// TIA Portal V19 export
FUNCTION_BLOCK "ULTRACHILLED_SKIDS"   // FB17, LAD
{ S7_Optimized_Access := 'TRUE' }
// stored: MemoryReserve 100, SetENOAutomatically false
   VAR_INPUT
      TEMP_SP : Real;
      START : Bool;
      STOP : Bool;
      AUTO : Bool;
      EMG : Bool;
      FS_HE_INLET : Bool;
      FS_HE_OUTLET : Bool;
      MGLT_LSP : Real;
      HOLD_RESUME : Bool;
      TT01_fault : Bool;
      TT02_fault : Bool;
      TT03_fault : Bool;
      TT04_fault : Bool;
      MGLT_FAULT : Bool;
      PUMP_1RPM : Real;
      "PUMP_1RPM SP" : Real;
      "PUMP_2 RPM" : Real;
      "PUMP_2 RPM SP" : Real;
      HEADER_PSP : Real;
      HEADER_PRESSURE_PV : Real;
      TEMP_PV : Real;
      MGLT_PV : Real;
   END_VAR
   VAR_OUTPUT
      PUMP_1_CMD : Bool;
      PUMP_2_CMD : Bool;
      RUNNING : Bool;
      UCH_BUXV1501_CMD : Bool;
      PUMP_1_FAULTY : Bool;
      PUMP_2_FAULTY : Bool;
   END_VAR
   VAR
      "STEP" : Int;
      ALL_OK : Bool;
      IEC_Timer_0_Instance { S7_SetPoint := 'True'} : TP_TIME;
      P_TRIG_1 { S7_SetPoint := 'True'} : Bool;
      P_TRIG_2 : Bool;
      P_TRIG_3 : Bool;
      P_TRIG_4 : Bool;
      P_TRIG_5 : Bool;
      P_TRIG_6 : Bool;
      P_TRIG_7 : Bool;
      P_TRIG_8 : Bool;
   END_VAR
   VAR_TEMP   // added for the SCL form of the ladder/FBD networks
      _w1 : Bool;
      _w2 : Bool;
      _w3 : Bool;
      _w4 : Bool;
   END_VAR
BEGIN

REGION Network 1: PRECHECK
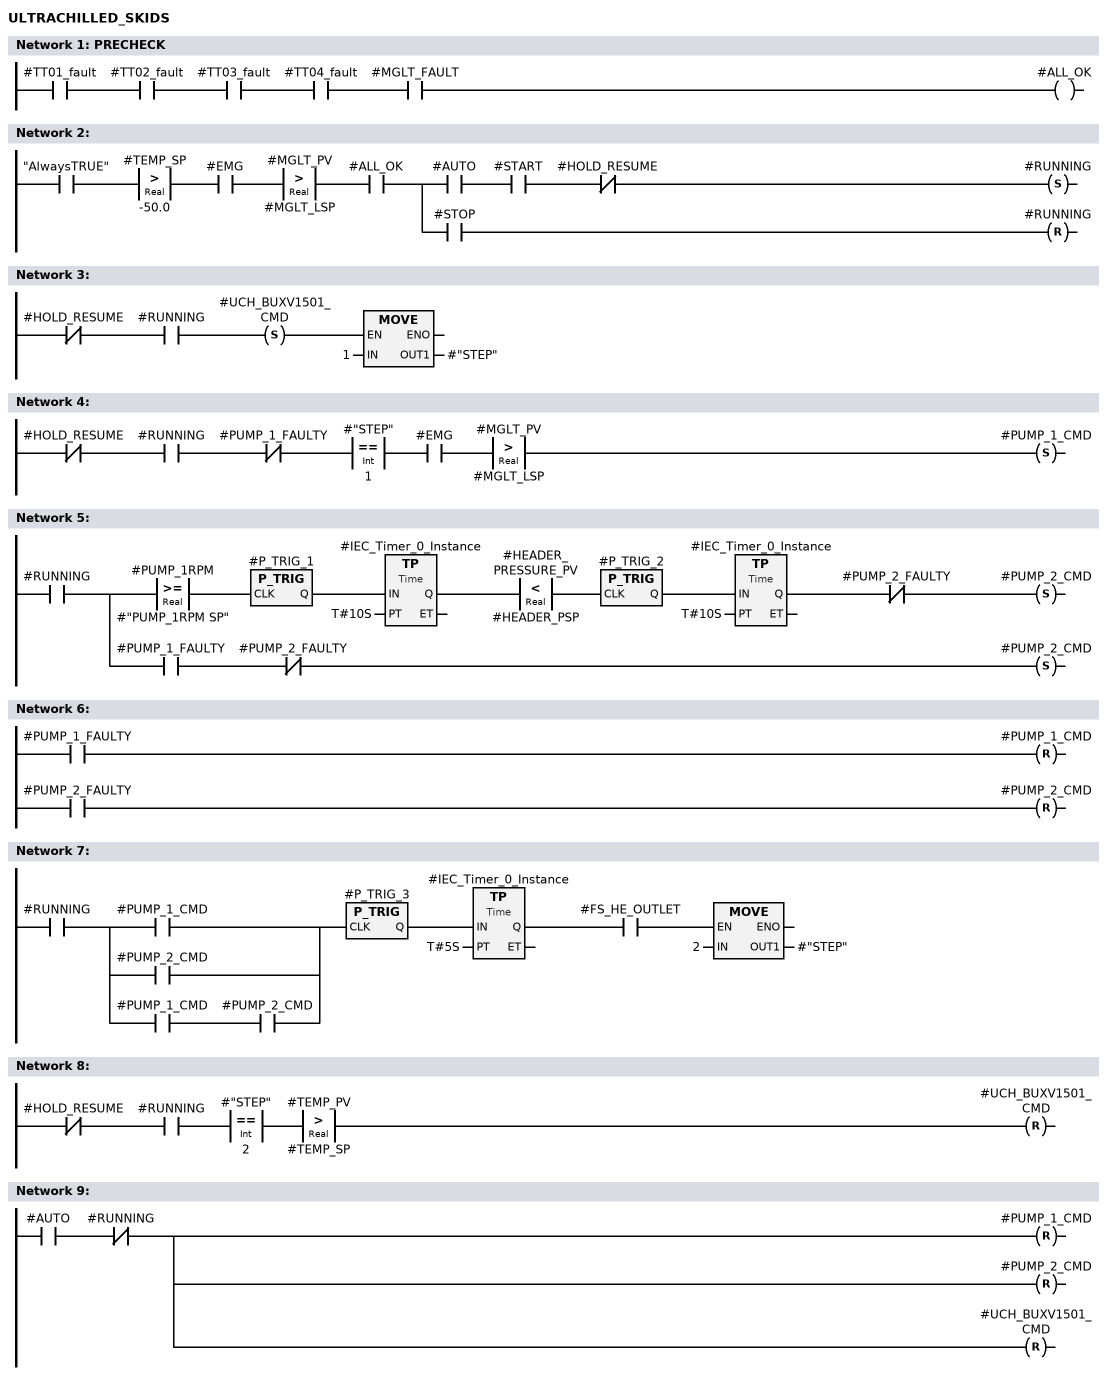
   RUNG wire#powerrail
      Contact( #TT01_fault )
      Contact( #TT02_fault )
      Contact( #TT03_fault )
      Contact( #TT04_fault )
      Contact( #MGLT_FAULT )
      Coil( #ALL_OK )
   END_RUNG
   // the same network as SCL:
   #ALL_OK := #TT01_fault AND #TT02_fault AND #TT03_fault AND #TT04_fault AND #MGLT_FAULT;
END_REGION

REGION Network 2
   RUNG wire#powerrail
      Contact( "AlwaysTRUE" )
      { S7_Templates := "SrcType := Real" } GT_Contact(in1 := #TEMP_SP, in2 := -50.0)
      Contact( #EMG )
      { S7_Templates := "SrcType := Real" } GT_Contact(in1 := #MGLT_PV, in2 := #MGLT_LSP)
      Contact( #ALL_OK )
      wire#w1
      Contact( #AUTO )
      Contact( #START )
      I_Contact( #HOLD_RESUME )
      S_Coil( #RUNNING )
   END_RUNG
   RUNG wire#w1
      Contact( #STOP )
      R_Coil( #RUNNING )
   END_RUNG
   // the same network as SCL:
   #_w1 := "AlwaysTRUE" AND (#TEMP_SP > (-50.0)) AND #EMG AND (#MGLT_PV > #MGLT_LSP) AND #ALL_OK;
   IF #_w1 AND #AUTO AND #START AND NOT #HOLD_RESUME THEN #RUNNING := TRUE; END_IF;
   IF #_w1 AND #STOP THEN #RUNNING := FALSE; END_IF;
END_REGION

REGION Network 3
   RUNG wire#powerrail
      I_Contact( #HOLD_RESUME )
      Contact( #RUNNING )
      S_Coil( #UCH_BUXV1501_CMD )
      Move(in := 1, out1 => #"STEP")
   END_RUNG
   // the same network as SCL:
   IF NOT #HOLD_RESUME AND #RUNNING THEN
       #UCH_BUXV1501_CMD := TRUE;
       #"STEP" := 1;
   END_IF;
END_REGION

REGION Network 4
   RUNG wire#powerrail
      I_Contact( #HOLD_RESUME )
      Contact( #RUNNING )
      I_Contact( #PUMP_1_FAULTY )
      { S7_Templates := "SrcType := Int" } EQ_Contact(in1 := #"STEP", in2 := 1)
      Contact( #EMG )
      { S7_Templates := "SrcType := Real" } GT_Contact(in1 := #MGLT_PV, in2 := #MGLT_LSP)
      S_Coil( #PUMP_1_CMD )
   END_RUNG
   // the same network as SCL:
   IF NOT #HOLD_RESUME AND #RUNNING AND NOT #PUMP_1_FAULTY AND (#"STEP" = 1) AND #EMG AND (#MGLT_PV > #MGLT_LSP) THEN
       #PUMP_1_CMD := TRUE;
   END_IF;
END_REGION

REGION Network 5
   RUNG wire#powerrail
      Contact( #RUNNING )
      wire#w1
      { S7_Templates := "SrcType := Real" } GE_Contact(in1 := #PUMP_1RPM, in2 := #"PUMP_1RPM SP")
      P_Trig( #P_TRIG_1 )
      { S7_Templates := "time_type := Time" } #IEC_Timer_0_Instance.TP(pt := T#10S, et =>)
      { S7_Templates := "SrcType := Real" } LT_Contact(in1 := #HEADER_PRESSURE_PV, in2 := #HEADER_PSP)
      P_Trig( #P_TRIG_2 )
      { S7_Templates := "time_type := Time" } #IEC_Timer_0_Instance.TP(pt := T#10S, et =>)
      I_Contact( #PUMP_2_FAULTY )
      S_Coil( #PUMP_2_CMD )
   END_RUNG
   RUNG wire#w1
      Contact( #PUMP_1_FAULTY )
      I_Contact( #PUMP_2_FAULTY )
      S_Coil( #PUMP_2_CMD )
   END_RUNG
   // the same network as SCL:
   #_w1 := #RUNNING AND (#PUMP_1RPM >= #"PUMP_1RPM SP");
   #_w2 := #_w1 AND NOT #P_TRIG_1;   // rising edge
   #P_TRIG_1 := #_w1;
   #IEC_Timer_0_Instance(IN := #_w2, PT := T#10S);   // TP
   #_w3 := #IEC_Timer_0_Instance.Q AND (#HEADER_PRESSURE_PV < #HEADER_PSP);
   #_w4 := #_w3 AND NOT #P_TRIG_2;   // rising edge
   #P_TRIG_2 := #_w3;
   #IEC_Timer_0_Instance(IN := #_w4, PT := T#10S);   // TP
   IF #IEC_Timer_0_Instance.Q AND NOT #PUMP_2_FAULTY THEN #PUMP_2_CMD := TRUE; END_IF;
   IF #RUNNING AND #PUMP_1_FAULTY AND NOT #PUMP_2_FAULTY THEN #PUMP_2_CMD := TRUE; END_IF;
END_REGION

REGION Network 6
   RUNG wire#powerrail
      Contact( #PUMP_1_FAULTY )
      R_Coil( #PUMP_1_CMD )
   END_RUNG
   RUNG wire#powerrail
      Contact( #PUMP_2_FAULTY )
      R_Coil( #PUMP_2_CMD )
   END_RUNG
   // the same network as SCL:
   IF #PUMP_1_FAULTY THEN #PUMP_1_CMD := FALSE; END_IF;
   IF #PUMP_2_FAULTY THEN #PUMP_2_CMD := FALSE; END_IF;
END_REGION

REGION Network 7
   RUNG wire#powerrail
      Contact( #RUNNING )
      wire#w1
      Contact( #PUMP_1_CMD )
      wire#w2
      P_Trig( #P_TRIG_3 )
      { S7_Templates := "time_type := Time" } #IEC_Timer_0_Instance.TP(pt := T#5S, et =>)
      Contact( #FS_HE_OUTLET )
      Move(in := 2, out1 => #"STEP")
   END_RUNG
   RUNG wire#w1
      Contact( #PUMP_2_CMD )
   END_RUNG wire#w2
   RUNG wire#w1
      Contact( #PUMP_1_CMD )
      Contact( #PUMP_2_CMD )
   END_RUNG wire#w2
   // the same network as SCL:
   #_w1 := #RUNNING AND (#PUMP_1_CMD OR #PUMP_2_CMD OR (#PUMP_1_CMD AND #PUMP_2_CMD));
   #_w2 := #_w1 AND NOT #P_TRIG_3;   // rising edge
   #P_TRIG_3 := #_w1;
   #IEC_Timer_0_Instance(IN := #_w2, PT := T#5S);   // TP
   IF #IEC_Timer_0_Instance.Q AND #FS_HE_OUTLET THEN #"STEP" := 2; END_IF;
END_REGION

REGION Network 8
   RUNG wire#powerrail
      I_Contact( #HOLD_RESUME )
      Contact( #RUNNING )
      { S7_Templates := "SrcType := Int" } EQ_Contact(in1 := #"STEP", in2 := 2)
      { S7_Templates := "SrcType := Real" } GT_Contact(in1 := #TEMP_PV, in2 := #TEMP_SP)
      R_Coil( #UCH_BUXV1501_CMD )
   END_RUNG
   // the same network as SCL:
   IF NOT #HOLD_RESUME AND #RUNNING AND (#"STEP" = 2) AND (#TEMP_PV > #TEMP_SP) THEN
       #UCH_BUXV1501_CMD := FALSE;
   END_IF;
END_REGION

REGION Network 9
   RUNG wire#powerrail
      Contact( #AUTO )
      I_Contact( #RUNNING )
      wire#w1
      R_Coil( #PUMP_1_CMD )
   END_RUNG
   RUNG wire#w1
      R_Coil( #PUMP_2_CMD )
   END_RUNG
   RUNG wire#w1
      R_Coil( #UCH_BUXV1501_CMD )
   END_RUNG
   // the same network as SCL:
   IF #AUTO AND NOT #RUNNING THEN
       #PUMP_1_CMD := FALSE;
       #PUMP_2_CMD := FALSE;
       #UCH_BUXV1501_CMD := FALSE;
   END_IF;
END_REGION
END_FUNCTION_BLOCK
